RoboDK station: Bench V1 cell v8.rdk

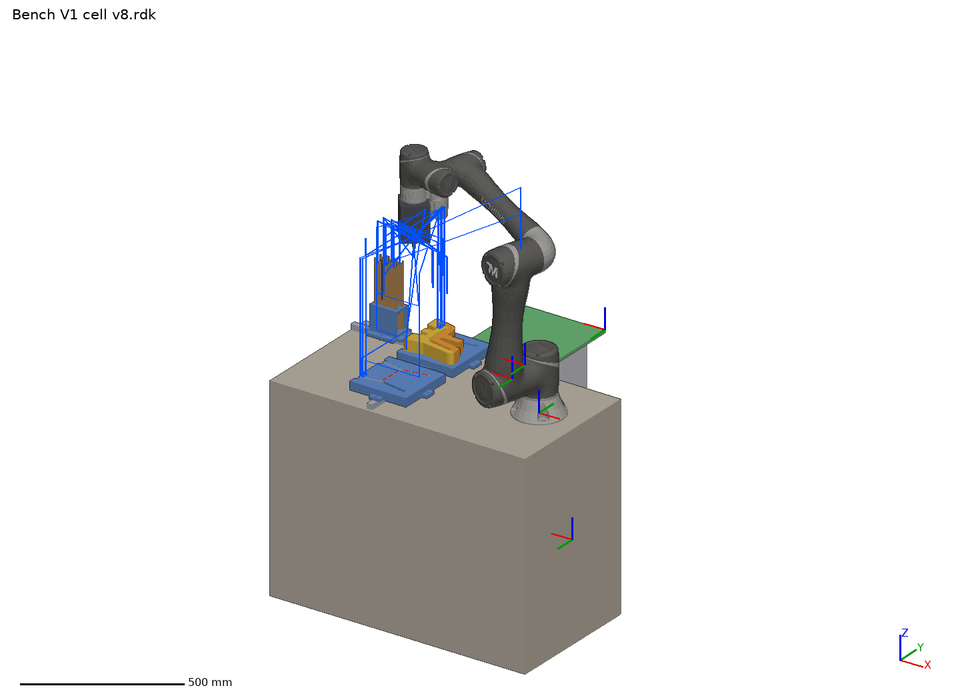
[picture v0: the station drawn from its stored meshes, robots at their saved joint values, targets as dots, program paths as lines]
Station Bench V1 cell v8 (saved by RoboDK 6.1.1). Poses are relative to the parent item; angles as X-Y-Z fixed-axis rotations.
  - frame Cell at (0, 0, 0) mm
    - frame Work plate at (-206.44, 152.99, -4.46) mm, rotated rx -0.03 ry -0.07 rz -179.98 deg
      - frame Ground base at (0, -67, 20) mm
        - object Table at (0, 0, 0) mm, size 950 x 510 x 730 mm
        - object Profile A-B at (0, 0, 0) mm, size 20 x 540 x 20 mm
        - object Profile rack at (0, 0, 0) mm, size 240 x 20 x 20 mm
        - object Base A at (235, 95, 10) mm, rotated rx 0 ry 0 rz 90 deg, size 246 x 246 x 32 mm, geometry from frame_jig_v8.stl
        - object Base B at (235, 345, 10) mm, rotated rx 0 ry 0 rz 90 deg, size 246 x 246 x 32 mm, geometry from frame_jig_v8.stl
        - object Plank jig at (420, 30, 0) mm, size 136 x 96 x 102 mm, geometry from plank_rack_v8.stl
        - frame AMR at (-60, -340, 0) mm
          - object AMR plate at (0, 0, 0) mm, size 300 x 320 x 10 mm
          - object AMR top module at (0, 0, 0) mm, size 220 x 240 x 377 mm
          - frame Omron LD-250 Base at (150, -40, -770) mm
            - robot AMR LD-250: 4 axes
                joint limits [-10000, -10000, -10, -3600] to [10000, 10000, 10, 3600]; home [0, 0, 0, 0]; saved at [0, 0, 0, 0]
        - object frame1 at (261.88, 92.28, 144.5) mm, size 174.7 x 141.9 x 10 mm, geometry from frame.stl
        - object frame2 at (261.88, 342.22, -95.5) mm, rotated rx -180 ry 0 rz 0 deg, size 174.7 x 141.9 x 10 mm, geometry from frame.stl
        - object piece A1 at (256.88, 92.28, 144.5) mm, rotated rx 90 ry 0 rz 90 deg, size 21.4 x 10 x 5 mm, geometry from interface_piece.stl
        - object piece B1 at (256.88, 342.22, 144.5) mm, rotated rx 90 ry 0 rz 90 deg, size 21.4 x 10 x 5 mm, geometry from interface_piece.stl
        - object plank1 at (435, 47.5, 128) mm, rotated rx 90 ry 0 rz 0 deg, size 25 x 250 x 5 mm, geometry from plank_body.stl
        - object piece A2 at (256.88, 62.3, 144.5) mm, rotated rx 90 ry 0 rz 90 deg, size 21.4 x 10 x 5 mm, geometry from interface_piece.stl
        - object piece B2 at (256.88, 372.2, 144.5) mm, rotated rx 90 ry 0 rz 90 deg, size 21.4 x 10 x 5 mm, geometry from interface_piece.stl
        - object plank2 at (465, 47.5, 128) mm, rotated rx 90 ry 0 rz 0 deg, size 25 x 250 x 5 mm, geometry from plank_body.stl
        - object piece A3 at (256.88, 122.27, 144.5) mm, rotated rx 90 ry 0 rz 90 deg, size 21.4 x 10 x 5 mm, geometry from interface_piece.stl
        - object piece B3 at (256.88, 312.23, 144.5) mm, rotated rx 90 ry 0 rz 90 deg, size 21.4 x 10 x 5 mm, geometry from interface_piece.stl
        - object plank3 at (495, 47.5, 128) mm, rotated rx 90 ry 0 rz 0 deg, size 25 x 250 x 5 mm, geometry from plank_body.stl
        - object piece A4 at (238.44, 144.24, 144.5) mm, rotated rx 90 ry 0 rz 170 deg, size 21.4 x 10 x 5 mm, geometry from interface_piece.stl
        - object piece B4 at (238.44, 290.26, 144.5) mm, rotated rx 90 ry 0 rz 10 deg, size 21.4 x 10 x 5 mm, geometry from interface_piece.stl
        - object plank4 at (435, 77.5, 128) mm, rotated rx 90 ry 0 rz 0 deg, size 25 x 250 x 5 mm, geometry from plank_body.stl
        - object piece A5 at (208.91, 149.45, 144.5) mm, rotated rx 90 ry 0 rz 170 deg, size 21.4 x 10 x 5 mm, geometry from interface_piece.stl
        - object piece B5 at (208.91, 285.05, 144.5) mm, rotated rx 90 ry 0 rz 10 deg, size 21.4 x 10 x 5 mm, geometry from interface_piece.stl
        - object plank5 at (465, 77.5, 128) mm, rotated rx 90 ry 0 rz 0 deg, size 25 x 250 x 5 mm, geometry from plank_body.stl
        - object piece A6 at (179.38, 154.66, 144.5) mm, rotated rx 90 ry 0 rz 170 deg, size 21.4 x 10 x 5 mm, geometry from interface_piece.stl
        - object piece B6 at (179.38, 279.84, 144.5) mm, rotated rx 90 ry 0 rz 10 deg, size 21.4 x 10 x 5 mm, geometry from interface_piece.stl
        - object plank6 at (495, 77.5, 128) mm, rotated rx 90 ry 0 rz 0 deg, size 25 x 250 x 5 mm, geometry from plank_body.stl
        - object Guide inner at (235, 95, 10) mm, rotated rx 0 ry 0 rz 90 deg, size 158.3 x 160 x 40 mm, geometry from guide_inner_v7.stl
        - object Guide outer at (235, 95, 10) mm, rotated rx 0 ry 0 rz 90 deg, size 177.7 x 180 x 40 mm, geometry from guide_outer_v7.stl
        - target Home (Cartesian target) at (260, 220, 380) mm, rotated rx 180 ry 0 rz 0 deg; joints [-15.175, 7.513, -83.536, -13.906, -90.009, 74.801] of Omron TM5-900
        - target plank3 pick travel (Cartesian target) at (495, 45, 380) mm, rotated rx 180 ry 0 rz -90 deg; joints [-23.734, -31.934, -35.025, -22.97, -89.998, 156.242] of Omron TM5-900
        - target plank3 pick approach (Cartesian target) at (495, 45, 278) mm, rotated rx 180 ry 0 rz -90 deg; joints [-23.733, -27.239, -56.964, -5.726, -89.998, 156.243] of Omron TM5-900
        - target plank3 pick (Cartesian target) at (495, 45, 238) mm, rotated rx 180 ry 0 rz -90 deg; joints [-23.733, -26.931, -63.004, 0.007, -89.998, 156.243] of Omron TM5-900
        - target plank3 pick out (Cartesian target) at (495, 45, 298) mm, rotated rx 180 ry 0 rz -90 deg; joints [-23.733, -27.648, -53.545, -8.735, -89.998, 156.243] of Omron TM5-900
        - target plank3 pick up (Cartesian target) at (495, 45, 380) mm, rotated rx 180 ry 0 rz -90 deg; joints [-23.734, -31.934, -35.025, -22.97, -89.998, 156.242] of Omron TM5-900
        - target plank3 place travel (Cartesian target) at (259.38, 122.27, 380) mm, rotated rx 180 ry 0 rz 0 deg; joints [-26.735, 6.228, -82.41, -13.747, -89.994, 63.241] of Omron TM5-900
        - target plank3 above guide (Cartesian target) at (259.38, 122.27, 329.5) mm, rotated rx 180 ry 0 rz 0 deg; joints [-26.734, 7.429, -90.62, -6.738, -89.994, 63.242] of Omron TM5-900
        - target plank3 place (Cartesian target) at (259.38, 122.27, 254.5) mm, rotated rx 180 ry 0 rz 0 deg; joints [-26.733, 7.696, -101.324, 3.699, -89.994, 63.243] of Omron TM5-900
        - target plank3 push approach (Cartesian target) at (259.38, 122.27, 289.5) mm, rotated rx 180 ry 0 rz 0 deg; joints [-26.734, 7.799, -96.531, -1.197, -89.994, 63.242] of Omron TM5-900
        - target plank3 push (Cartesian target) at (259.38, 122.27, 269.5) mm, rotated rx 180 ry 0 rz 0 deg; joints [-26.734, 7.79, -99.311, 1.592, -89.994, 63.242] of Omron TM5-900
        - target plank3 push out (Cartesian target) at (259.38, 122.27, 289.5) mm, rotated rx 180 ry 0 rz 0 deg; joints [-26.734, 7.799, -96.531, -1.197, -89.994, 63.242] of Omron TM5-900
        - target plank3 place up (Cartesian target) at (259.38, 122.27, 380) mm, rotated rx 180 ry 0 rz 0 deg; joints [-26.735, 6.228, -82.41, -13.747, -89.994, 63.241] of Omron TM5-900
        - target plank6 pick travel (Cartesian target) at (495, 75, 380) mm, rotated rx 180 ry 0 rz -90 deg; joints [-21.493, -30.518, -37.272, -22.138, -90.001, 158.482] of Omron TM5-900
        - target plank6 pick approach (Cartesian target) at (495, 75, 278) mm, rotated rx 180 ry 0 rz -90 deg; joints [-21.494, -26.175, -58.531, -5.222, -90.001, 158.482] of Omron TM5-900
        - target plank6 pick (Cartesian target) at (495, 75, 238) mm, rotated rx 180 ry 0 rz -90 deg; joints [-21.494, -25.923, -64.482, 0.477, -90.001, 158.482] of Omron TM5-900
        - target plank6 pick out (Cartesian target) at (495, 75, 298) mm, rotated rx 180 ry 0 rz -90 deg; joints [-21.494, -26.548, -55.176, -8.204, -90.001, 158.482] of Omron TM5-900
        - target plank6 pick up (Cartesian target) at (495, 75, 380) mm, rotated rx 180 ry 0 rz -90 deg; joints [-21.493, -30.518, -37.272, -22.138, -90.001, 158.482] of Omron TM5-900
        - target plank6 place travel (Cartesian target) at (179.82, 157.12, 380) mm, rotated rx 180 ry 0 rz 80 deg; joints [-27.46, 17.648, -91.296, -16.281, -89.993, -17.484] of Omron TM5-900
        - target plank6 above guide (Cartesian target) at (179.82, 157.12, 329.5) mm, rotated rx 180 ry 0 rz 80 deg; joints [-27.459, 19.163, -99.527, -9.564, -89.993, -17.483] of Omron TM5-900
        - target plank6 place (Cartesian target) at (179.82, 157.12, 254.5) mm, rotated rx 180 ry 0 rz 80 deg; joints [-27.458, 19.968, -110.552, 0.655, -89.993, -17.482] of Omron TM5-900
        - target plank6 push approach (Cartesian target) at (179.82, 157.12, 289.5) mm, rotated rx 180 ry 0 rz 80 deg; joints [-27.459, 19.817, -105.571, -4.174, -89.993, -17.483] of Omron TM5-900
        - target plank6 push (Cartesian target) at (179.82, 157.12, 269.5) mm, rotated rx 180 ry 0 rz 80 deg; joints [-27.458, 19.954, -108.451, -1.431, -89.993, -17.482] of Omron TM5-900
        - target plank6 push out (Cartesian target) at (179.82, 157.12, 289.5) mm, rotated rx 180 ry 0 rz 80 deg; joints [-27.459, 19.817, -105.571, -4.174, -89.993, -17.483] of Omron TM5-900
        - target plank6 place up (Cartesian target) at (179.82, 157.12, 380) mm, rotated rx 180 ry 0 rz 80 deg; joints [-27.46, 17.648, -91.296, -16.281, -89.993, -17.484] of Omron TM5-900
        - target plank2 pick travel (Cartesian target) at (465, 45, 380) mm, rotated rx 180 ry 0 rz -90 deg; joints [-24.747, -26.16, -43.947, -19.821, -89.997, 155.229] of Omron TM5-900
        - target plank2 pick approach (Cartesian target) at (465, 45, 278) mm, rotated rx 180 ry 0 rz -90 deg; joints [-24.747, -22.712, -63.497, -3.719, -89.997, 155.229] of Omron TM5-900
        - target plank2 pick (Cartesian target) at (465, 45, 238) mm, rotated rx 180 ry 0 rz -90 deg; joints [-24.747, -22.62, -69.206, 1.897, -89.997, 155.229] of Omron TM5-900
        - target plank2 pick out (Cartesian target) at (465, 45, 298) mm, rotated rx 180 ry 0 rz -90 deg; joints [-24.747, -22.985, -60.313, -6.63, -89.997, 155.229] of Omron TM5-900
        - target plank2 pick up (Cartesian target) at (465, 45, 380) mm, rotated rx 180 ry 0 rz -90 deg; joints [-24.747, -26.16, -43.947, -19.821, -89.997, 155.229] of Omron TM5-900
        - target plank2 place travel (Cartesian target) at (259.38, 62.3, 380) mm, rotated rx 180 ry 0 rz 0 deg; joints [-33.11, 4.08, -80.465, -13.545, -89.986, 56.866] of Omron TM5-900
        - target plank2 above guide (Cartesian target) at (259.38, 62.3, 329.5) mm, rotated rx 180 ry 0 rz 0 deg; joints [-33.109, 5.258, -88.697, -6.491, -89.986, 56.867] of Omron TM5-900
        - target plank2 place (Cartesian target) at (259.38, 62.3, 254.5) mm, rotated rx 180 ry 0 rz 0 deg; joints [-33.106, 5.48, -99.369, 3.96, -89.986, 56.87] of Omron TM5-900
        - target plank2 push approach (Cartesian target) at (259.38, 62.3, 289.5) mm, rotated rx 180 ry 0 rz 0 deg; joints [-33.107, 5.604, -94.599, -0.935, -89.986, 56.869] of Omron TM5-900
        - target plank2 push (Cartesian target) at (259.38, 62.3, 269.5) mm, rotated rx 180 ry 0 rz 0 deg; joints [-33.107, 5.582, -97.368, 1.856, -89.986, 56.869] of Omron TM5-900
        - target plank2 push out (Cartesian target) at (259.38, 62.3, 289.5) mm, rotated rx 180 ry 0 rz 0 deg; joints [-33.107, 5.604, -94.599, -0.935, -89.986, 56.869] of Omron TM5-900
        - target plank2 place up (Cartesian target) at (259.38, 62.3, 380) mm, rotated rx 180 ry 0 rz 0 deg; joints [-33.11, 4.08, -80.465, -13.545, -89.986, 56.866] of Omron TM5-900
        - target plank5 pick travel (Cartesian target) at (465, 75, 380) mm, rotated rx 180 ry 0 rz -90 deg; joints [-22.426, -24.899, -45.812, -19.217, -90, 157.55] of Omron TM5-900
        - target plank5 pick approach (Cartesian target) at (465, 75, 278) mm, rotated rx 180 ry 0 rz -90 deg; joints [-22.426, -21.667, -64.958, -3.304, -90, 157.55] of Omron TM5-900
        - target plank5 pick (Cartesian target) at (465, 75, 238) mm, rotated rx 180 ry 0 rz -90 deg; joints [-22.426, -21.616, -70.607, 2.294, -90, 157.55] of Omron TM5-900
        - target plank5 pick out (Cartesian target) at (465, 75, 298) mm, rotated rx 180 ry 0 rz -90 deg; joints [-22.426, -21.914, -61.816, -6.199, -90, 157.55] of Omron TM5-900
        - target plank5 pick up (Cartesian target) at (465, 75, 380) mm, rotated rx 180 ry 0 rz -90 deg; joints [-22.426, -24.899, -45.812, -19.217, -90, 157.55] of Omron TM5-900
        - target plank5 place travel (Cartesian target) at (209.34, 151.91, 380) mm, rotated rx 180 ry 0 rz 80 deg; joints [-26.173, 13.604, -88.427, -15.105, -89.995, -16.197] of Omron TM5-900
        - target plank5 above guide (Cartesian target) at (209.34, 151.91, 329.5) mm, rotated rx 180 ry 0 rz 80 deg; joints [-26.172, 14.971, -96.63, -8.269, -89.995, -16.196] of Omron TM5-900
        - target plank5 place (Cartesian target) at (209.34, 151.91, 254.5) mm, rotated rx 180 ry 0 rz 80 deg; joints [-26.171, 15.525, -107.517, 2.064, -89.995, -16.195] of Omron TM5-900
        - target plank5 push approach (Cartesian target) at (209.34, 151.91, 289.5) mm, rotated rx 180 ry 0 rz 80 deg; joints [-26.172, 15.494, -102.614, -2.808, -89.995, -16.196] of Omron TM5-900
        - target plank5 push (Cartesian target) at (209.34, 151.91, 269.5) mm, rotated rx 180 ry 0 rz 80 deg; joints [-26.171, 15.562, -105.452, -0.038, -89.995, -16.195] of Omron TM5-900
        - target plank5 push out (Cartesian target) at (209.34, 151.91, 289.5) mm, rotated rx 180 ry 0 rz 80 deg; joints [-26.172, 15.494, -102.614, -2.808, -89.995, -16.196] of Omron TM5-900
        - target plank5 place up (Cartesian target) at (209.34, 151.91, 380) mm, rotated rx 180 ry 0 rz 80 deg; joints [-26.173, 13.604, -88.427, -15.105, -89.995, -16.197] of Omron TM5-900
        - target plank1 pick travel (Cartesian target) at (435, 45, 380) mm, rotated rx 180 ry 0 rz -90 deg; joints [-25.849, -21.109, -51.235, -17.585, -89.995, 154.127] of Omron TM5-900
        - target plank1 pick approach (Cartesian target) at (435, 45, 278) mm, rotated rx 180 ry 0 rz -90 deg; joints [-25.848, -18.423, -69.366, -2.14, -89.995, 154.128] of Omron TM5-900
        - target plank1 pick (Cartesian target) at (435, 45, 238) mm, rotated rx 180 ry 0 rz -90 deg; joints [-25.848, -18.485, -74.861, 3.418, -89.995, 154.128] of Omron TM5-900
        - target plank1 pick out (Cartesian target) at (435, 45, 298) mm, rotated rx 180 ry 0 rz -90 deg; joints [-25.848, -18.602, -66.333, -4.993, -89.995, 154.128] of Omron TM5-900
        - target plank1 pick up (Cartesian target) at (435, 45, 380) mm, rotated rx 180 ry 0 rz -90 deg; joints [-25.849, -21.109, -51.235, -17.585, -89.995, 154.127] of Omron TM5-900
        - target plank1 place travel (Cartesian target) at (259.38, 92.28, 380) mm, rotated rx 180 ry 0 rz 0 deg; joints [-30.002, 5.273, -81.555, -13.646, -89.99, 59.974] of Omron TM5-900
        - target plank1 above guide (Cartesian target) at (259.38, 92.28, 329.5) mm, rotated rx 180 ry 0 rz 0 deg; joints [-30.001, 6.462, -89.773, -6.618, -89.99, 59.975] of Omron TM5-900
        - target plank1 place (Cartesian target) at (259.38, 92.28, 254.5) mm, rotated rx 180 ry 0 rz 0 deg; joints [-29.999, 6.707, -100.462, 3.826, -89.99, 59.977] of Omron TM5-900
        - target plank1 push approach (Cartesian target) at (259.38, 92.28, 289.5) mm, rotated rx 180 ry 0 rz 0 deg; joints [-30, 6.82, -95.68, -1.07, -89.99, 59.976] of Omron TM5-900
        - target plank1 push (Cartesian target) at (259.38, 92.28, 269.5) mm, rotated rx 180 ry 0 rz 0 deg; joints [-29.999, 6.805, -98.455, 1.721, -89.99, 59.977] of Omron TM5-900
        - target plank1 push out (Cartesian target) at (259.38, 92.28, 289.5) mm, rotated rx 180 ry 0 rz 0 deg; joints [-30, 6.82, -95.68, -1.07, -89.99, 59.976] of Omron TM5-900
        - target plank1 place up (Cartesian target) at (259.38, 92.28, 380) mm, rotated rx 180 ry 0 rz 0 deg; joints [-30.002, 5.273, -81.555, -13.646, -89.99, 59.974] of Omron TM5-900
        - target plank4 pick travel (Cartesian target) at (435, 75, 380) mm, rotated rx 180 ry 0 rz -90 deg; joints [-23.442, -19.915, -52.889, -17.125, -89.998, 156.534] of Omron TM5-900
        - target plank4 pick approach (Cartesian target) at (435, 75, 278) mm, rotated rx 180 ry 0 rz -90 deg; joints [-23.441, -17.374, -70.754, -1.801, -89.998, 156.534] of Omron TM5-900
        - target plank4 pick (Cartesian target) at (435, 75, 238) mm, rotated rx 180 ry 0 rz -90 deg; joints [-23.441, -17.469, -76.208, 3.749, -89.998, 156.535] of Omron TM5-900
        - target plank4 pick out (Cartesian target) at (435, 75, 298) mm, rotated rx 180 ry 0 rz -90 deg; joints [-23.441, -17.535, -67.75, -4.644, -89.998, 156.534] of Omron TM5-900
        - target plank4 pick up (Cartesian target) at (435, 75, 380) mm, rotated rx 180 ry 0 rz -90 deg; joints [-23.442, -19.915, -52.889, -17.125, -89.998, 156.534] of Omron TM5-900
        - target plank4 place travel (Cartesian target) at (238.87, 146.7, 380) mm, rotated rx 180 ry 0 rz 80 deg; joints [-25.064, 9.56, -85.255, -14.234, -89.996, -15.088] of Omron TM5-900
        - target plank4 above guide (Cartesian target) at (238.87, 146.7, 329.5) mm, rotated rx 180 ry 0 rz 80 deg; joints [-25.064, 10.82, -93.45, -7.299, -89.996, -15.088] of Omron TM5-900
        - target plank4 place (Cartesian target) at (238.87, 146.7, 254.5) mm, rotated rx 180 ry 0 rz 80 deg; joints [-25.063, 11.191, -104.224, 3.105, -89.996, -15.087] of Omron TM5-900
        - target plank4 push approach (Cartesian target) at (238.87, 146.7, 289.5) mm, rotated rx 180 ry 0 rz 80 deg; joints [-25.063, 11.246, -99.387, -1.787, -89.996, -15.088] of Omron TM5-900
        - target plank4 push (Cartesian target) at (238.87, 146.7, 269.5) mm, rotated rx 180 ry 0 rz 80 deg; joints [-25.063, 11.265, -102.19, 0.997, -89.996, -15.087] of Omron TM5-900
        - target plank4 push out (Cartesian target) at (238.87, 146.7, 289.5) mm, rotated rx 180 ry 0 rz 80 deg; joints [-25.063, 11.246, -99.387, -1.787, -89.996, -15.088] of Omron TM5-900
        - target plank4 place up (Cartesian target) at (238.87, 146.7, 380) mm, rotated rx 180 ry 0 rz 80 deg; joints [-25.064, 9.56, -85.255, -14.234, -89.996, -15.088] of Omron TM5-900
        - target guide A-B pick out low (Cartesian target) at (305, -2, 50) mm, rotated rx 0 ry -90 rz -90 deg; joints [-54.001, -55.302, -66.544, -58.121, -54.025, -90.047] of Omron TM5-900
        - target guide A-B pick out (Cartesian target) at (305, -2, 450) mm, rotated rx 0 ry -90 rz -90 deg; joints [-54.023, -46.797, -24.224, -108.946, -54.047, -90.047] of Omron TM5-900
        - target guide A-B via (Cartesian target) at (260, 220, 450) mm, rotated rx 0 ry -90 rz -90 deg; joints [-43.519, -15.63, -72.409, -91.922, -43.543, -90.038] of Omron TM5-900
        - target guide A-B pick (Cartesian target) at (305, 23, 50) mm, rotated rx 0 ry -90 rz -90 deg; joints [-52.769, -53.202, -70.764, -56, -52.793, -90.046] of Omron TM5-900
        - target guide A-B lift (Cartesian target) at (305, 23, 70) mm, rotated rx 0 ry -90 rz -90 deg; joints [-52.77, -51.654, -70.512, -57.8, -52.795, -90.046] of Omron TM5-900
        - target guide A-B up (Cartesian target) at (305, 23, 450) mm, rotated rx 0 ry -90 rz -90 deg; joints [-52.791, -42.108, -32.502, -105.356, -52.815, -90.046] of Omron TM5-900
        - target guide A-B across (Cartesian target) at (305, 411.5, 450) mm, rotated rx 0 ry -90 rz -90 deg; joints [-22.822, -12.347, -76.526, -91.058, -22.846, -90.002] of Omron TM5-900
        - target guide A-B place (Cartesian target) at (305, 411.5, 50) mm, rotated rx 0 ry 90 rz -90 deg; joints [32.16, -52.809, -71.628, -55.614, -147.864, 90.109] of Omron TM5-900
        - target guide A-B half turned (Cartesian target) at (305, 411.5, 510) mm, rotated rx 180 ry 0 rz 90 deg; joints [7.658, -11.756, -43.444, -34.738, -90.036, 7.634] of Omron TM5-900
        - target guide A-B over place (Cartesian target) at (305, 411.5, 450) mm, rotated rx 0 ry 90 rz -90 deg; joints [32.194, -41.276, -33.995, -104.779, -147.83, 90.109] of Omron TM5-900
        - target guide A-B place approach (Cartesian target) at (305, 411.5, 90) mm, rotated rx 0 ry 90 rz -90 deg; joints [32.164, -49.767, -70.99, -59.293, -147.86, 90.109] of Omron TM5-900
        - target guide A-B place out (Cartesian target) at (305, 436.5, 50) mm, rotated rx 0 ry 90 rz -90 deg; joints [33.903, -54.873, -67.483, -57.693, -146.121, 90.107] of Omron TM5-900
        - target guide A-B place out up (Cartesian target) at (305, 436.5, 450) mm, rotated rx 0 ry 90 rz -90 deg; joints [33.937, -45.706, -26.251, -108.092, -146.087, 90.107] of Omron TM5-900
        - target sub pick (Cartesian target) at (331.7, 155.8, 22) mm, rotated rx -120 ry 0 rz 99.93 deg; joints [-10.817, -49.592, -62.944, -35.703, -107.89, -10.723] of Omron TM5-900
        - target sub pick approach (Cartesian target) at (331.7, 155.8, 62) mm, rotated rx -120 ry 0 rz 99.93 deg; joints [-10.816, -47.47, -60.886, -39.884, -107.889, -10.723] of Omron TM5-900
        - target sub via (Cartesian target) at (260, 220, 450) mm, rotated rx -120 ry 0 rz 99.93 deg; joints [-6.662, -47.029, -4.332, -97.506, -104.344, -8.467] of Omron TM5-900
        - target sub to middle (joint target) at (235, 220, 450) mm, rotated rx -120 ry 0 rz 99.93 deg; joints [-6.912, -35.827, -24.869, -88.137, -104.559, -8.601] of Omron TM5-900
        - target sub place (Cartesian target) at (331.7, 278.7, 267) mm, rotated rx 60 ry 0 rz -99.93 deg; joints [-7.772, -66.43, -63.352, 99.835, 88.147, -1.05] of Omron TM5-900
        - target sub wrist ready (Cartesian target) at (235, 220, 450) mm, rotated rx -97.05 ry -56.07 rz -41.34 deg; joints [-61.447, 21.783, -105.714, -80.63, -14.785, -41.381] of Omron TM5-900
        - target sub wrist swapped (joint target) at (299.46, 101.48, 487.12) mm, rotated rx -83.11 ry -56.1 rz -81.48 deg; joints [-61.447, 21.783, -105.714, -80.63, 14.785, -41.381] of Omron TM5-900
        - target sub above guide (Cartesian target) at (331.7, 278.7, 342) mm, rotated rx 60 ry 0 rz -99.93 deg; joints [-7.771, -59.69, -64.836, 94.579, 88.145, -1.051] of Omron TM5-900
        - target sub flipped high (Cartesian target) at (331.7, 278.7, 450) mm, rotated rx 60 ry 0 rz -99.93 deg; joints [-7.768, -51.697, -63.403, 85.153, 88.143, -1.052] of Omron TM5-900
        - target sub flipped (Cartesian target) at (331.7, 278.7, 387) mm, rotated rx 60 ry 0 rz -99.93 deg; joints [-7.77, -56.096, -64.751, 90.9, 88.144, -1.051] of Omron TM5-900
        - target sub place out (Cartesian target) at (353.03, 274.97, 254.5) mm, rotated rx 60 ry 0 rz -99.93 deg; joints [-7.832, -70.217, -57.092, 97.363, 88.198, -1.02] of Omron TM5-900
        - target sub clear (Cartesian target) at (203.03, 274.97, 254.5) mm, rotated rx 60 ry 0 rz -99.93 deg; joints [-9.686, -55.841, -91.233, 117.144, 89.805, -0.095] of Omron TM5-900
        - target sub back to middle (Cartesian target) at (260, 220, 450) mm, rotated rx 60 ry 0 rz -99.93 deg; joints [-13.363, -42.859, -79.991, 92.875, 92.991, 1.741] of Omron TM5-900
        - target inner pick out low (Cartesian target) at (300, 436.5, 50) mm, rotated rx 0 ry 90 rz -90 deg; joints [34.133, -54.429, -68.375, -57.244, -145.891, 90.106] of Omron TM5-900
        - target inner pick out (Cartesian target) at (300, 436.5, 450) mm, rotated rx 0 ry 90 rz -90 deg; joints [34.167, -44.687, -28.062, -107.299, -145.857, 90.106] of Omron TM5-900
        - target inner via (Cartesian target) at (260, 220, 450) mm, rotated rx 0 ry 90 rz -90 deg; joints [17.44, -15.684, -72.376, -92.03, -162.584, 90.152] of Omron TM5-900
        - target inner centre (Cartesian target) at (260, 220, 450) mm, rotated rx 60 ry 0 rz -99.93 deg; joints [-13.363, -42.859, -79.991, 92.875, 92.991, 1.741] of Omron TM5-900
        - target inner wrist ready (Cartesian target) at (260, 220, 450) mm, rotated rx 84.7 ry -42.38 rz 141.25 deg; joints [-56.29, 6.341, -129.876, 107.647, 14.521, 27.028] of Omron TM5-900
        - target inner wrist swapped (joint target) at (333.3, 109.99, 412.23) mm, rotated rx 95.4 ry -42.35 rz 106.06 deg; joints [-56.29, 6.341, -129.876, 107.647, -14.521, 27.028] of Omron TM5-900
        - target inner via (Cartesian target) at (260, 220, 450) mm, rotated rx 0 ry 90 rz -90 deg; joints [17.44, -15.684, -72.376, -92.03, -162.584, 90.152] of Omron TM5-900
        - target inner pick (Cartesian target) at (300, 411.5, 50) mm, rotated rx 0 ry 90 rz -90 deg; joints [32.385, -52.376, -72.498, -55.177, -147.639, 90.109] of Omron TM5-900
        - target inner out 1 (Cartesian target) at (298.61, 419.38, 50) mm, rotated rx 0 ry 90 rz -90 deg; joints [33.008, -52.886, -71.474, -55.689, -147.016, 90.108] of Omron TM5-900
        - target inner out 2 (Cartesian target) at (298.61, 419.38, 100) mm, rotated rx 0 ry 90 rz -90 deg; joints [33.013, -49.136, -70.588, -60.325, -147.012, 90.108] of Omron TM5-900
        - target inner out 3 (Cartesian target) at (98.61, 419.38, 100) mm, rotated rx 0 ry 90 rz -90 deg; joints [44.708, -34.806, -97.302, -47.93, -135.316, 90.094] of Omron TM5-900
        - target inner up (Cartesian target) at (98.61, 419.38, 450) mm, rotated rx 0 ry 90 rz -90 deg; joints [44.75, -18.939, -68.149, -92.951, -135.274, 90.094] of Omron TM5-900
        - target inner across (Cartesian target) at (300, 23, 450) mm, rotated rx 0 ry 90 rz -90 deg; joints [-5.115, -18.297, -99.746, 118.345, -174.861, 269.767] of Omron TM5-900
        - target inner place (Cartesian target) at (300, 23, 50) mm, rotated rx 0 ry -90 rz -90 deg; joints [-53.104, -52.768, -71.637, -55.562, -53.128, 269.954] of Omron TM5-900
        - target inner over place (Cartesian target) at (300, 23, 450) mm, rotated rx 0 ry -90 rz -90 deg; joints [-53.126, -41.231, -34.01, -104.725, -53.15, 269.954] of Omron TM5-900
        - target inner place approach (Cartesian target) at (300, 23, 90) mm, rotated rx 0 ry -90 rz -90 deg; joints [-53.107, -49.726, -70.999, -59.242, -53.131, 269.954] of Omron TM5-900
        - target inner place out (Cartesian target) at (300, -2, 50) mm, rotated rx 0 ry -90 rz -90 deg; joints [-54.333, -54.855, -67.442, -57.67, -54.357, 269.953] of Omron TM5-900
        - target inner place out up (Cartesian target) at (300, -2, 450) mm, rotated rx 0 ry -90 rz -90 deg; joints [-54.355, -45.716, -26.165, -108.085, -54.379, 269.953] of Omron TM5-900
        - target outer pick out low (Cartesian target) at (310, 436.5, 50) mm, rotated rx 0 ry 90 rz -90 deg; joints [33.675, -55.323, -66.576, -58.15, -146.349, 90.107] of Omron TM5-900
        - target outer pick out (Cartesian target) at (310, 436.5, 450) mm, rotated rx 0 ry 90 rz -90 deg; joints [33.709, -46.795, -24.294, -108.959, -146.315, 90.107] of Omron TM5-900
        - target outer via (Cartesian target) at (260, 220, 450) mm, rotated rx 0 ry 90 rz -90 deg; joints [17.44, -15.684, -72.376, -92.03, -162.584, 90.152] of Omron TM5-900
        - target outer pick (Cartesian target) at (310, 411.5, 50) mm, rotated rx 0 ry 90 rz -90 deg; joints [31.938, -53.247, -70.746, -56.058, -148.086, 90.11] of Omron TM5-900
        - target outer out 1 (Cartesian target) at (318, 411.5, 50) mm, rotated rx 0 ry 90 rz -90 deg; joints [31.587, -53.963, -69.306, -56.782, -148.437, 90.11] of Omron TM5-900
        - target outer out 2 (Cartesian target) at (318, 411.5, 100) mm, rotated rx 0 ry 90 rz -90 deg; joints [31.591, -50.274, -68.409, -61.369, -148.433, 90.11] of Omron TM5-900
        - target outer out 3 (Cartesian target) at (318, 226.5, 100) mm, rotated rx 0 ry 90 rz -90 deg; joints [16.316, -38.054, -91.333, -50.709, -163.708, 90.159] of Omron TM5-900
        - target outer out 4 (Cartesian target) at (393, 226.5, 100) mm, rotated rx 0 ry 90 rz -90 deg; joints [14.468, -45.46, -77.534, -57.114, -165.557, 90.171] of Omron TM5-900
        - target outer up (Cartesian target) at (393, 226.5, 450) mm, rotated rx 0 ry 90 rz -90 deg; joints [14.491, -35.028, -44.344, -100.735, -165.534, 90.171] of Omron TM5-900
        - target outer across (Cartesian target) at (310, 23, 450) mm, rotated rx 0 ry 90 rz -90 deg; joints [-5.014, -19.515, -98.061, 117.883, -174.962, 269.761] of Omron TM5-900
        - target outer place (Cartesian target) at (310, 23, 50) mm, rotated rx 0 ry -90 rz -90 deg; joints [-52.438, -53.643, -69.877, -56.446, -52.462, 269.954] of Omron TM5-900
        - target outer over place (Cartesian target) at (310, 23, 450) mm, rotated rx 0 ry -90 rz -90 deg; joints [-52.459, -43.023, -30.914, -106.028, -52.483, 269.954] of Omron TM5-900
        - target outer place approach (Cartesian target) at (310, 23, 90) mm, rotated rx 0 ry -90 rz -90 deg; joints [-52.44, -50.641, -69.232, -60.093, -52.464, 269.954] of Omron TM5-900
        - target outer place out (Cartesian target) at (310, -2, 50) mm, rotated rx 0 ry -90 rz -90 deg; joints [-53.672, -55.755, -65.631, -58.58, -53.697, 269.953] of Omron TM5-900
        - target outer place out up (Cartesian target) at (310, -2, 450) mm, rotated rx 0 ry -90 rz -90 deg; joints [-53.694, -47.966, -22.101, -109.899, -53.718, 269.953] of Omron TM5-900
        - target bench pick out low (Cartesian target) at (331.7, 278.7, 287) mm, rotated rx 180 ry 0 rz -99.93 deg; joints [-6.796, -1.217, -88.401, -0.313, -90.019, 183.106] of Omron TM5-900
        - target bench pick out (Cartesian target) at (331.7, 278.7, 322) mm, rotated rx 180 ry 0 rz -99.93 deg; joints [-6.795, -1.443, -83.283, -5.205, -90.019, 183.108] of Omron TM5-900
        - target bench via (Cartesian target) at (260, 220, 450) mm, rotated rx 180 ry 0 rz -99.93 deg; joints [-15.173, 4.405, -70.453, -23.881, -90.009, 174.729] of Omron TM5-900
        - target bench pick (Cartesian target) at (331.7, 278.7, 262) mm, rotated rx 180 ry 0 rz -99.93 deg; joints [-6.797, -1.3, -91.802, 3.172, -90.019, 183.105] of Omron TM5-900
        - target bench lift (Cartesian target) at (331.7, 278.7, 362) mm, rotated rx 180 ry 0 rz -99.93 deg; joints [-6.793, -2.201, -76.864, -10.866, -90.019, 183.109] of Omron TM5-900
        - target bench over AMR (Cartesian target) at (186.7, -246.3, 362) mm, rotated rx 180 ry 0 rz -99.93 deg; joints [-61.468, -11.92, -65.859, -12.166, -89.954, 128.434] of Omron TM5-900
        - target bench down (Cartesian target) at (186.7, -246.3, 243) mm, rotated rx 180 ry 0 rz -99.93 deg; joints [-61.459, -10.857, -83.828, 4.741, -89.954, 128.443] of Omron TM5-900
        - target bench place out (Cartesian target) at (186.7, -246.3, 283) mm, rotated rx 180 ry 0 rz -99.93 deg; joints [-61.462, -10.67, -78.47, -0.805, -89.954, 128.44] of Omron TM5-900
        - target bench place out up (Cartesian target) at (186.7, -246.3, 450) mm, rotated rx 180 ry 0 rz -99.93 deg; joints [-61.475, -16.59, -46.875, -26.479, -89.954, 128.428] of Omron TM5-900
        - target back to middle (Cartesian target) at (260, 220, 450) mm, rotated rx -180 ry 0 rz -99.93 deg; joints [-15.173, 4.405, -70.453, -23.881, -90.009, 174.729] of Omron TM5-900
    - frame Omron TM5-900 Base at (0, 0, 0) mm
      - robot Omron TM5-900: 6 axes, payload 4 kg, reach 900 mm, repeatability 0.05 mm, weight 22.6 kg
          modified DH rows (alpha deg, a mm, theta deg, d mm): 0, 0, 0, 145.2; 90, 0, 90, 0; 0, 429, 0, 0; 0, 411, -90, 122.3; -90, 0, 0, 106.5; 90, 0, 180, 114.15
          joint limits [-270, -180, -155, -180, -180, -270] to [270, 180, 155, 180, 180, 270]; home [0, 0, 90, -90, 90, 0]; saved at [-15.174, 6.177, -77.285, -18.821, -90.009, 124.765]
        - tool EGP, TCP at (0, 0, 160) mm, size 94 x 90 x 160 mm
  - program AssembleBench (324 instructions, listed below)
  - Python program Deliver (AMR) (listed below)
  - Python program Assemble and deliver (listed below)
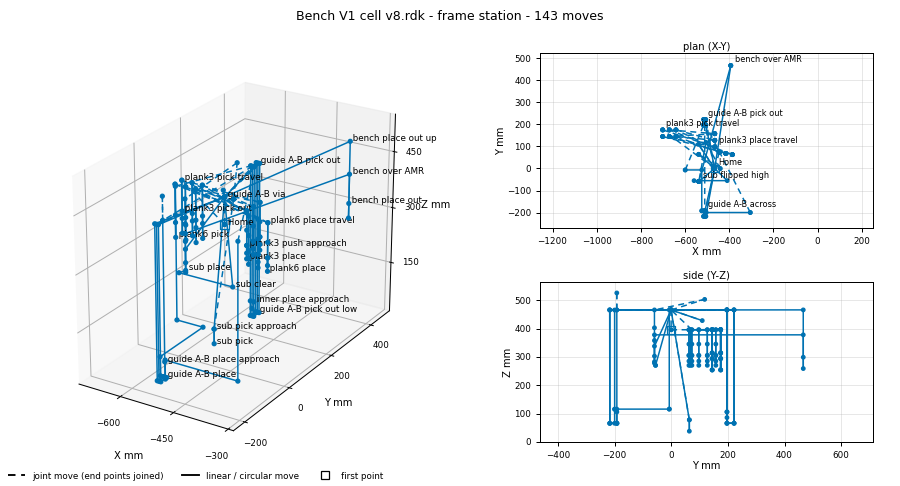
[picture p0: tool path of Bench V1 cell v8.rdk in frame station, 143 of 143 moves have a stored position in this frame; points joined in program order, loops and branches not executed]

--- program AssembleBench (robot Omron TM5-900) ---
  Simulation: parts to start
  Set Ref.: Ground base
  Set Tool: EGP
  Smooth(0)
  Set speed (100.0 mm/s)
  MoveJ (Home)
  MoveJ (plank3 pick travel)
  MoveL (plank3 pick approach)
  Set speed (20.0 mm/s)
  MoveL (plank3 pick)
  Set IO_0=1
  Pause 500 ms
  Simulation: attach plank3
  MoveL (plank3 pick out)
  Set speed (100.0 mm/s)
  MoveL (plank3 pick up)
  MoveJ (plank3 place travel)
  MoveL (plank3 above guide)
  Set speed (20.0 mm/s)
  MoveL (plank3 place)
  Set IO_0=0
  Pause 500 ms
  Simulation: release plank3
  MoveL (plank3 push approach)
  Set IO_0=1
  Pause 300 ms
  MoveL (plank3 push)
  MoveL (plank3 push out)
  Set IO_0=0
  Pause 300 ms
  Set speed (100.0 mm/s)
  MoveL (plank3 place up)
  MoveJ (plank6 pick travel)
  MoveL (plank6 pick approach)
  Set speed (20.0 mm/s)
  MoveL (plank6 pick)
  Set IO_0=1
  Pause 500 ms
  Simulation: attach plank6
  MoveL (plank6 pick out)
  Set speed (100.0 mm/s)
  MoveL (plank6 pick up)
  MoveJ (plank6 place travel)
  MoveL (plank6 above guide)
  Set speed (20.0 mm/s)
  MoveL (plank6 place)
  Set IO_0=0
  Pause 500 ms
  Simulation: release plank6
  MoveL (plank6 push approach)
  Set IO_0=1
  Pause 300 ms
  MoveL (plank6 push)
  MoveL (plank6 push out)
  Set IO_0=0
  Pause 300 ms
  Set speed (100.0 mm/s)
  MoveL (plank6 place up)
  MoveJ (plank2 pick travel)
  MoveL (plank2 pick approach)
  Set speed (20.0 mm/s)
  MoveL (plank2 pick)
  Set IO_0=1
  Pause 500 ms
  Simulation: attach plank2
  MoveL (plank2 pick out)
  Set speed (100.0 mm/s)
  MoveL (plank2 pick up)
  MoveJ (plank2 place travel)
  MoveL (plank2 above guide)
  Set speed (20.0 mm/s)
  MoveL (plank2 place)
  Set IO_0=0
  Pause 500 ms
  Simulation: release plank2
  MoveL (plank2 push approach)
  Set IO_0=1
  Pause 300 ms
  MoveL (plank2 push)
  MoveL (plank2 push out)
  Set IO_0=0
  Pause 300 ms
  Set speed (100.0 mm/s)
  MoveL (plank2 place up)
  MoveJ (plank5 pick travel)
  MoveL (plank5 pick approach)
  Set speed (20.0 mm/s)
  MoveL (plank5 pick)
  Set IO_0=1
  Pause 500 ms
  Simulation: attach plank5
  MoveL (plank5 pick out)
  Set speed (100.0 mm/s)
  MoveL (plank5 pick up)
  MoveJ (plank5 place travel)
  MoveL (plank5 above guide)
  Set speed (20.0 mm/s)
  MoveL (plank5 place)
  Set IO_0=0
  Pause 500 ms
  Simulation: release plank5
  MoveL (plank5 push approach)
  Set IO_0=1
  Pause 300 ms
  MoveL (plank5 push)
  MoveL (plank5 push out)
  Set IO_0=0
  Pause 300 ms
  Set speed (100.0 mm/s)
  MoveL (plank5 place up)
  MoveJ (plank1 pick travel)
  MoveL (plank1 pick approach)
  Set speed (20.0 mm/s)
  MoveL (plank1 pick)
  Set IO_0=1
  Pause 500 ms
  Simulation: attach plank1
  MoveL (plank1 pick out)
  Set speed (100.0 mm/s)
  MoveL (plank1 pick up)
  MoveJ (plank1 place travel)
  MoveL (plank1 above guide)
  Set speed (20.0 mm/s)
  MoveL (plank1 place)
  Set IO_0=0
  Pause 500 ms
  Simulation: release plank1
  MoveL (plank1 push approach)
  Set IO_0=1
  Pause 300 ms
  MoveL (plank1 push)
  MoveL (plank1 push out)
  Set IO_0=0
  Pause 300 ms
  Set speed (100.0 mm/s)
  MoveL (plank1 place up)
  MoveJ (plank4 pick travel)
  MoveL (plank4 pick approach)
  Set speed (20.0 mm/s)
  MoveL (plank4 pick)
  Set IO_0=1
  Pause 500 ms
  Simulation: attach plank4
  MoveL (plank4 pick out)
  Set speed (100.0 mm/s)
  MoveL (plank4 pick up)
  MoveJ (plank4 place travel)
  MoveL (plank4 above guide)
  Set speed (20.0 mm/s)
  MoveL (plank4 place)
  Set IO_0=0
  Pause 500 ms
  Simulation: release plank4
  MoveL (plank4 push approach)
  Set IO_0=1
  Pause 300 ms
  MoveL (plank4 push)
  MoveL (plank4 push out)
  Set IO_0=0
  Pause 300 ms
  Set speed (100.0 mm/s)
  MoveL (plank4 place up)
  MoveJ (guide A-B via)
  MoveL (guide A-B pick out)
  MoveL (guide A-B pick out low)
  Set speed (20.0 mm/s)
  Set IO_0=1
  Pause 300 ms
  MoveL (guide A-B pick)
  Set IO_0=0
  Pause 500 ms
  Simulation: attach Guide inner
  Simulation: attach Guide outer
  MoveL (guide A-B lift)
  Set speed (100.0 mm/s)
  MoveL (guide A-B up)
  MoveJ (guide A-B across)
  MoveJ (guide A-B half turned)
  MoveJ (guide A-B over place)
  MoveL (guide A-B place approach)
  Set speed (20.0 mm/s)
  MoveL (guide A-B place)
  Set IO_0=1
  Pause 500 ms
  Simulation: release guide A-B
  MoveL (guide A-B place out)
  Set speed (100.0 mm/s)
  MoveL (guide A-B place out up)
  MoveJ (sub via)
  MoveL (sub pick approach)
  Set speed (20.0 mm/s)
  MoveL (sub pick)
  Set IO_0=1
  Pause 500 ms
  Simulation: attach frame1
  Simulation: attach plank1
  Simulation: attach plank2
  Simulation: attach plank3
  Simulation: attach plank4
  Simulation: attach plank5
  Simulation: attach plank6
  Simulation: attach piece A1
  Simulation: attach piece A2
  Simulation: attach piece A3
  Simulation: attach piece A4
  Simulation: attach piece A5
  Simulation: attach piece A6
  MoveL (sub pick approach)
  Set speed (100.0 mm/s)
  MoveJ (sub to middle)
  MoveL (sub wrist ready)
  MoveJ (sub wrist swapped)
  MoveJ (sub flipped high)
  MoveL (sub flipped)
  MoveL (sub above guide)
  Set speed (20.0 mm/s)
  MoveL (sub place)
  Set IO_0=0
  Pause 500 ms
  Simulation: release frame 1 with the planks
  MoveL (sub place out)
  MoveL (sub clear)
  MoveL (sub back to middle)
  Set speed (100.0 mm/s)
  MoveJ (inner centre)
  MoveL (inner wrist ready)
  MoveJ (inner wrist swapped)
  MoveL (inner via)
  MoveL (inner pick out)
  MoveL (inner pick out low)
  Set speed (20.0 mm/s)
  Set IO_0=1
  Pause 300 ms
  MoveL (inner pick)
  Set IO_0=0
  Pause 500 ms
  Simulation: attach Guide inner
  Set speed (20.0 mm/s)
  MoveL (inner out 1)
  MoveL (inner out 2)
  MoveL (inner out 3)
  Set speed (100.0 mm/s)
  MoveL (inner up)
  MoveJ (inner across)
  MoveJ (inner over place)
  MoveL (inner place approach)
  Set speed (20.0 mm/s)
  MoveL (inner place)
  Set IO_0=1
  Pause 500 ms
  Simulation: release inner
  MoveL (inner place out)
  Set speed (100.0 mm/s)
  MoveL (inner place out up)
  MoveJ (outer via)
  MoveL (outer pick out)
  MoveL (outer pick out low)
  Set speed (20.0 mm/s)
  Set IO_0=1
  Pause 300 ms
  MoveL (outer pick)
  Set IO_0=0
  Pause 500 ms
  Simulation: attach Guide outer
  Set speed (20.0 mm/s)
  MoveL (outer out 1)
  MoveL (outer out 2)
  MoveL (outer out 3)
  MoveL (outer out 4)
  Set speed (100.0 mm/s)
  MoveL (outer up)
  MoveJ (outer across)
  MoveJ (outer over place)
  MoveL (outer place approach)
  Set speed (20.0 mm/s)
  MoveL (outer place)
  Set IO_0=1
  Pause 500 ms
  Simulation: release outer
  MoveL (outer place out)
  Set speed (100.0 mm/s)
  MoveL (outer place out up)
  MoveJ (bench via)
  MoveL (bench pick out)
  MoveL (bench pick out low)
  Set speed (20.0 mm/s)
  Set IO_0=0
  Pause 300 ms
  MoveL (bench pick)
  Set IO_0=1
  Pause 500 ms
  Simulation: attach frame1
  Simulation: attach frame2
  Simulation: attach plank1
  Simulation: attach plank2
  Simulation: attach plank3
  Simulation: attach plank4
  Simulation: attach plank5
  Simulation: attach plank6
  Simulation: attach piece A1
  Simulation: attach piece A2
  Simulation: attach piece A3
  Simulation: attach piece A4
  Simulation: attach piece A5
  Simulation: attach piece A6
  Simulation: attach piece B1
  Simulation: attach piece B2
  Simulation: attach piece B3
  Simulation: attach piece B4
  Simulation: attach piece B5
  Simulation: attach piece B6
  MoveL (bench lift)
  Set speed (100.0 mm/s)
  MoveL (bench over AMR)
  Set speed (20.0 mm/s)
  MoveL (bench down)
  Set IO_0=0
  Pause 500 ms
  Simulation: release bench
  MoveL (bench place out)
  Set speed (100.0 mm/s)
  MoveL (bench place out up)
  MoveL (back to middle)
  MoveJ (Home)

--- Python program Deliver (AMR) ---
"""The AMR drives the finished bench 2 m away along the table and comes back (RoboDK station script
"Deliver (AMR)").

    python robot_cell/amr_drive.py           also works from outside RoboDK

Needs only the robodk package. Everything under the station's "AMR" frame rides along: its plate,
top module and LD-250, and the bench once the robot program has set it down there (the program's
release puts the bench under the AMR frame).
"""
import time

from robodk import robolink, robomath

DISTANCE = 2000          # mm, along the ground base's x (away from the robot)
STEPS = 120              # per direction
PAUSE = 1.0              # s at the far end
OWN = ("AMR plate", "AMR top module")


def main():
    RDK = robolink.Robolink()
    amr = RDK.Item("AMR", robolink.ITEM_TYPE_FRAME)
    if not amr.Valid():
        raise SystemExit("no AMR in the open station")
    riding = [c for c in amr.Childs() if c.Type() == robolink.ITEM_TYPE_OBJECT and c.Name() not in OWN]
    home = amr.Pose()
    for out in (True, False):
        for i in range(1, STEPS + 1):
            s = i / STEPS if out else 1 - i / STEPS
            s = 0.5 - 0.5 * robomath.cos(robomath.pi * s)        # smooth start and stop
            amr.setPose(robomath.transl(DISTANCE * s, 0, 0) * home)
            RDK.Render(True)
            time.sleep(0.02)
        if out:
            time.sleep(PAUSE)
    amr.setPose(home)
    print(f"AMR drove {DISTANCE / 1000:.0f} m and back with {len(riding)} parts on its plate")


if __name__ == "__main__":
    main()

--- Python program Assemble and deliver ---
"""The whole cycle (station script "Assemble and deliver"): the robot program AssembleBench builds the
bench and sets it down on the AMR, then the AMR drives it 2 m along the table and back (amr_drive.py).

    python robot_cell/assemble_and_deliver.py      also works from outside RoboDK
"""
import time

from robodk import robolink

import amr_drive


def main():
    RDK = robolink.Robolink()
    prog = RDK.Item("AssembleBench", robolink.ITEM_TYPE_PROGRAM)
    if not prog.Valid():
        raise SystemExit("no AssembleBench in the open station")
    t0 = time.time()
    prog.RunProgram()
    time.sleep(1)
    while prog.Busy():
        time.sleep(0.2)
    print(f"AssembleBench done after {time.time() - t0:.0f} s (at the simulation speed)")
    amr_drive.main()


if __name__ == "__main__":
    main()
